FUNCTION_BLOCK FB_Besturing IMPLEMENTS ITF_Besturing
VAR_INPUT
END_VAR
VAR_OUTPUT
END_VAR
VAR
END_VAR

{warning 'Add method implementation '}
METHOD StatusLampGeel : BOOL
END_METHOD

{warning 'Add method implementation '}
METHOD StatusLampGroen : BOOL
END_METHOD

{warning 'Add method implementation '}
METHOD StatusLampRood : BOOL
END_METHOD

END_FUNCTION_BLOCK

(* stored: Version 1.1.0.1
   POU FB_Besturing: Id {2d50245b-8b53-4c5f-a24c-67422698d9cd}, SpecialFunc None
   Folder Methods: Id {cbf70383-cc63-4fb1-bda0-6b79f4aa4a91}
   Method StatusLampGeel: Id {6fdd2845-507c-4f65-969d-037b60785eaa}
   Method StatusLampGroen: Id {1ae9ab3f-ab41-464b-ae60-e994a85e5dbc}
   Method StatusLampRood: Id {9ad9db52-d671-4976-8c61-563214ae33a3} *)
